SYSTEM epuck_functionblocks
  (* Standard: 61499-2; Classification: Application; ApplicationDomain: Robotics; Function: Simulation; Type: Application; Description: Function blocks network for the epuck1 robot routine *)
  (* Version 1.0, 2026-10-22, Mauricio Martins Taques Filho, GASR/UDESC, Initial version *)
  APPLICATION epuck_functionblocksApp
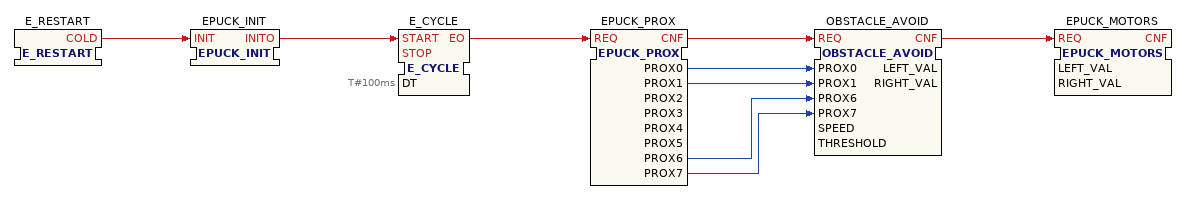
    FBS
      E_CYCLE : E_CYCLE(DT := T#100ms);
      E_RESTART : E_RESTART;
      EPUCK_PROX : EPUCK_PROX;
      EPUCK_MOTORS : EPUCK_MOTORS;
      EPUCK_INIT : EPUCK_INIT;
      OBSTACLE_AVOID : OBSTACLE_AVOID;
    END_FBS
    EVENT_CONNECTIONS
      E_RESTART.COLD TO EPUCK_INIT.INIT;
      EPUCK_INIT.INITO TO E_CYCLE.START;
      E_CYCLE.EO TO EPUCK_PROX.REQ;
      OBSTACLE_AVOID.CNF TO EPUCK_MOTORS.REQ;
      EPUCK_PROX.CNF TO OBSTACLE_AVOID.REQ;
    END_CONNECTIONS
    DATA_CONNECTIONS
      EPUCK_PROX.PROX0 TO OBSTACLE_AVOID.PROX0;
      EPUCK_PROX.PROX1 TO OBSTACLE_AVOID.PROX1;
      EPUCK_PROX.PROX6 TO OBSTACLE_AVOID.PROX6;
      EPUCK_PROX.PROX7 TO OBSTACLE_AVOID.PROX7;
    END_CONNECTIONS
  END_APPLICATION
END_SYSTEM
